(* IEC 61131-3 sources: SRCI_CLIENT_PLC/RobotLibrary/Library/POUs/Trigger/MC_WaitTime/Structures, 4 files *)

(* ---- WaitTimeOutCmd.st ---- *)
{attribute 'pack_mode' := '1'}
// -------------------------------------------------------------------------
//  SRCI Robot Library
// -------------------------------------------------------------------------
//
//  Object:      WaitTimeOutCmd
//  Author:      Thorsten Brach
//  Date:        2024-06-30
//
//  Description:
//
//
//  Copyright:
//    (C) 2024 Thorsten Brach. All rights reserved
//             Licensed under the MIT License.
//
//  Disclaimer:
//    This project is provided without any guarantee and can be used for
//    private and commercial purposes. Any use is at the user’s
//    own risk and responsibility.
//
// -------------------------------------------------------------------------
TYPE WaitTimeOutCmd :
STRUCT
  /// Current value of time [ms] that has elapsed since processing of the command has started.
  ElapsedTime        : UDINT;
END_STRUCT
END_TYPE

(* ---- WaitTimeParCmd.st ---- *)
{attribute 'pack_mode' := '1'}
// -------------------------------------------------------------------------
//  SRCI Robot Library
// -------------------------------------------------------------------------
//
//  Object:      WaitTimeParCmd
//  Author:      Thorsten Brach
//  Date:        2024-06-30
//
//  Description:
//
//
//  Copyright:
//    (C) 2024 Thorsten Brach. All rights reserved
//             Licensed under the MIT License.
//
//  Disclaimer:
//    This project is provided without any guarantee and can be used for
//    private and commercial purposes. Any use is at the user’s
//    own risk and responsibility.
//
// -------------------------------------------------------------------------
TYPE WaitTimeParCmd :
STRUCT
  /// Duration [ms] of the waiting time. The value of the parameter must be positive
  WaitTime           : UDINT;
END_STRUCT
END_TYPE

(* ---- WaitTimeRecvData.st ---- *)
{attribute 'pack_mode' := '1'}
// -------------------------------------------------------------------------
//  SRCI Robot Library
// -------------------------------------------------------------------------
//
//  Object:      WaitTimeRecvData
//  Author:      Thorsten Brach
//  Date:        2024-06-30
//
//  Description:
//
//
//  Copyright:
//    (C) 2024 Thorsten Brach. All rights reserved
//             Licensed under the MIT License.
//
//  Disclaimer:
//    This project is provided without any guarantee and can be used for
//    private and commercial purposes. Any use is at the user’s
//    own risk and responsibility.
//
// -------------------------------------------------------------------------
TYPE WaitTimeRecvData EXTENDS RspHeader :
STRUCT
  /// Current value of time [ms] that has elapsed since processing of the command has started.
  ElapsedTime : UDINT;
  /// Reserve
  Reserve1    : BYTE;
  /// Reserve
  Reserve2    : BYTE;
  /// Reserve
  Reserve3    : BYTE;
  /// Reserve
  Reserve4    : BYTE;
END_STRUCT
END_TYPE

(* ---- WaitTimeSendData.st ---- *)
{attribute 'pack_mode' := '1'}
// -------------------------------------------------------------------------
//  SRCI Robot Library
// -------------------------------------------------------------------------
//
//  Object:      WaitTimeSendData
//  Author:      Thorsten Brach
//  Date:        2024-06-30
//
//  Description:
//
//
//  Copyright:
//    (C) 2024 Thorsten Brach. All rights reserved
//             Licensed under the MIT License.
//
//  Disclaimer:
//    This project is provided without any guarantee and can be used for
//    private and commercial purposes. Any use is at the user’s
//    own risk and responsibility.
//
// -------------------------------------------------------------------------
TYPE WaitTimeSendData EXTENDS CmdHeader:
STRUCT
  /// Duration [ms] of the waiting time. The value of the parameter must be positive
  WaitTime : UDINT;
  /// Reserve
  Reserve1 : BYTE;
  /// Reserve
  Reserve2 : BYTE;
  /// Reserve
  Reserve3 : BYTE;
  /// Reserve
  Reserve4 : BYTE;
END_STRUCT
END_TYPE
